FUNCTION_BLOCK Test_AssertEquals_STRING EXTENDS T_UnitTestBase IMPLEMENTS I_UnitTest
VAR

END_VAR

{attribute 'analysis' := '-33'} // inhibit unused variable warning
METHOD RunTest
VAR
    Expected : T_MaxString := 'A long string,A long string,A long string,A long string,A long string,A long string,A long string,A long string,A long string,A long string,A long string,A long string';
    Actual   : T_MaxString := 'A very long string,A long string,A long string,A long string,A long string,A long string,A long string,A long string,A long string,A long string,A long string,A long string';
END_VAR
THIS^.AssertEquals_STRING(Expected := Expected,
                          Actual   := Actual,
                          Message  := 'Assertion is not working correctly');

						  
// Should fail the assertion!
						  
TestCompleted();
END_METHOD

END_FUNCTION_BLOCK

(* stored: Version 1.1.0.1, ProductVersion 3.1.4026.19
   POU Test_AssertEquals_STRING: Id {75079ee0-e49c-438a-aaa2-185999de7306}, SpecialFunc None
   Method RunTest: Id {f4bcfeff-7dbf-4d88-90f0-b5bec5ba1bd0} *)
